Fanuc KAREL source: KA00191.KL

PROGRAM KA00191
%NOLOCKGROUP
VAR
  SRC: ARRAY[4] OF SHORT
  DST: ARRAY[4] OF REAL
BEGIN
  DST = SRC
END KA00191
